(* IEC 61131-3 sources: cds-text-sync-reference-project/project-view/CODESYS_Linux_SL/PLC Logic/CI_CD_Application/GVL, 1 file *)

(* ---- GVL_Test.st ---- *)
VAR_GLOBAL
	// Test flags for CI/CD
	g_xTestSuiteRunning : BOOL := FALSE;
	g_xAllPassed : BOOL := FALSE;
	g_uiTestCount : UINT := 0;
	g_uiPassCount : UINT := 0;
	g_uiFailCount : UINT := 0;
END_VAR
